PROGRAM Control_FBD
VAR
	
	ixPulse			AT %I*:	BOOL; 		(* PULS button *)
	ixStart			AT %I*:	BOOL; 		(* START switch *)
	ixSetLevel		AT %I*:	BOOL; 		(* NIVÅ switch *)
	ixLevel3		AT %I*:	BOOL; 		(* Sensor for level 3 *)
	ixLevel2		AT %I*:	BOOL; 		(* Sensor for level 2 *)
	ixLevel1		AT %I*:	BOOL; 		(* Sensor for level 1 *)
	ixNotEmpty		AT %I*:	BOOL; 		(* Sensor for not empty *)
	ixTempOk		AT %I*:	BOOL; 		(* Temp sensor *)
	
	mxFill : BOOL;
	mxForw : BOOL;
	mxBack : BOOL;
	mxSpin : BOOL;
	mxDrain : BOOL;
	mxHeat : BOOL;
	
	qxForw			AT %Q*:	BOOL; 		(* Washer cylinder forward *)
	qxBack			AT %Q*:	BOOL; 		(* Washer cylinder back *)
	qxSpin			AT %Q*:	BOOL; 		(* Hi-spin/Centrifuge need qxForw or qxBack*)
	qxFill			AT %Q*:	BOOL; 		(* Fill water *)
	qxDrain			AT %Q*:	BOOL; 		(* Drain water *)
	qxHeat			AT %Q*:	BOOL; 		(* Heat water *)
	qxDispBit1		AT %Q*:	BOOL; 		(* Display bit 1 *)
	qxDispBit2		AT %Q*:	BOOL; 		(* Display bit 2 *)
END_VAR

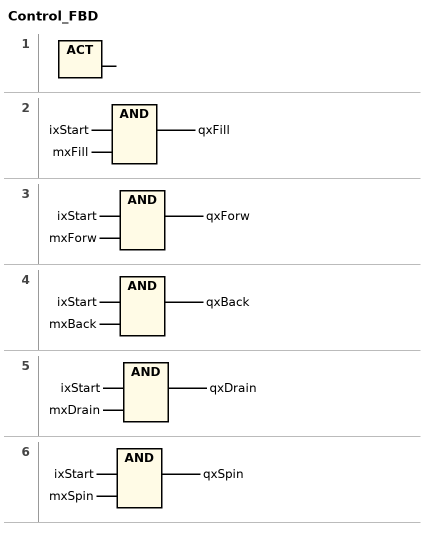
// NETWORK 1
ACT();

// NETWORK 2
qxFill := ixStart AND mxFill;

// NETWORK 3
qxForw := ixStart AND mxForw;

// NETWORK 4
qxBack := ixStart AND mxBack;

// NETWORK 5
qxDrain := ixStart AND mxDrain;

// NETWORK 6
qxSpin := ixStart AND mxSpin;

ACTION ACT:
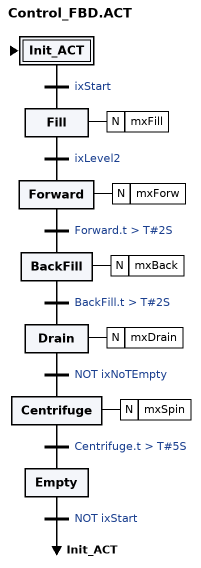
INITIAL_STEP Init_ACT:
END_STEP
TRANSITION FROM Init_ACT TO Fill
    := ixStart;
END_TRANSITION
STEP Fill:
    mxFill(N);
END_STEP
TRANSITION FROM Fill TO Forward
    := ixLevel2;
END_TRANSITION
STEP Forward:
    mxForw(N);
END_STEP
TRANSITION FROM Forward TO BackFill
    := Forward.t > T#2S;
END_TRANSITION
STEP BackFill:
    mxBack(N);
END_STEP
TRANSITION FROM BackFill TO Drain
    := BackFill.t > T#2S;
END_TRANSITION
STEP Drain:
    mxDrain(N);
END_STEP
TRANSITION FROM Drain TO Centrifuge
    := NOT ixNoTEmpty;
END_TRANSITION
STEP Centrifuge:
    mxSpin(N);
END_STEP
TRANSITION FROM Centrifuge TO Empty
    := Centrifuge.t > T#5S;
END_TRANSITION
STEP Empty:
END_STEP
TRANSITION FROM Empty TO Init_ACT
    := NOT ixStart;
END_TRANSITION
END_ACTION

END_PROGRAM

(* stored: Version 1.1.0.1
   POU Control_FBD: Id {84d3f40d-a0f6-423e-bc58-eeabb716185d}, SpecialFunc None
   Action ACT: Id {45b4c563-5046-4a28-bdc8-7e9e98e1e4a0} *)
